(* IEC 61131-3 sources: codesys-to-s7/tests/corpus/C2S7-SEM-TEMP/pos, 1 file *)

(* ---- input.st ---- *)
FUNCTION_BLOCK FB_Case
VAR
    a : INT;
END_VAR
VAR_TEMP
    tmp : INT;
END_VAR
a := tmp + 1;
END_FUNCTION_BLOCK
